{attribute 'no_assign'}
FUNCTION_BLOCK FB_DO_WTURBINE_LD0_WCNV1_Torq EXTENDS FB_AcsiCommonDataClass
VAR_INPUT
	mag: FB_AcsiDATypeAnalogueValue := (Fc:=ACSI_FC_MX, TrgOp:=ACSI_TrgOp_dchg OR ACSI_TrgOp_dupd, i:=(bPresence:=FALSE), bLinkResult:=THIS^.AddDataToContainer(ipData:=mag));
	q: FB_AcsiDATypeQuality := (Fc:=ACSI_FC_MX, TrgOp:=ACSI_TrgOp_qchg, bLinkResult:=THIS^.AddDataToContainer(ipData:=q));
	t: FB_AcsiDATypeTimeStamp := (Fc:=ACSI_FC_MX, bLinkResult:=THIS^.AddDataToContainer(ipData:=t));
END_VAR
VAR
END_VAR

END_FUNCTION_BLOCK

(* stored: Version 1.1.0.1
   POU FB_DO_WTURBINE_LD0_WCNV1_Torq: Id {bfb1e473-e238-4e18-bd9f-31289cffdfb2}, SpecialFunc None *)
